Fanuc KAREL source: KA00004.KL

PROGRAM KA00004
%NOLOCKGROUP
VAR
  SRC: INTEGER
  DST: STRING[80]
BEGIN
  SRC = 2
  DST = SRC
END KA00004
